// TIA Portal V20 export
// export: Created 2026-10-11T05:19:06.4640986Z, ExportSetting WithDefaults, DisplayName Totally Integrated Automation Portal, DisplayVersion V20, DisplayName TIA Portal Openness, DisplayVersion V20, DisplayName TIA Portal Teamcenter Gateway, DisplayVersion V20, DisplayName TIA Portal Version Control Interface, DisplayVersion V20, DisplayName SINAMICS Startdrive Advanced, DisplayVersion V20 SP1 Update 2, DisplayName SINAMICS Startdrive G110M, G120, G120C, G120D, G120P, G115D, DisplayVersion V20 SP1 Update 2, DisplayName SINAMICS Startdrive G130, G150, S120, S150, SINAMICS MV, G220, S200, S210, DisplayVersion V20 SP1 Update 2, DisplayName STEP 7 Professional, DisplayVersion V20, DisplayName STEP 7 Safety, DisplayVersion V20, DisplayName WinCC Basic/Comfort/Advanced, DisplayVersion V20, DisplayName WinCC Professional, DisplayVersion V20, DisplayName WinCC Unified, DisplayVersion V20
FUNCTION "FRK_Route_InnerUnit" : Bool   // FC65, SCL
{ S7_Optimized_Access := 'TRUE' }
VERSION : 0.1
// stored: AutoNumber true, IsIECCheckEnabled false, SetENOAutomatically false, UDAEnableTagReadback false
   VAR_INPUT
      Request : "ST_HmiRequest";
   END_VAR
   VAR_IN_OUT
      Module : "FB_InnerUnit";
      Hal : "ST_InnerUnitHal";
      Report : "ST_ReleaseReport";
   END_VAR
   VAR_TEMP
      RouteMatched : Bool;
      Index : Int;
   END_VAR
BEGIN

   #FRK_Route_InnerUnit := FALSE;
   IF NOT "FRK_PathOwned"(OwnerPath := #Module.Status.Name, TargetPath := #Request.TargetPath) THEN
       RETURN;
   END_IF;
   "FRK_Release_InnerUnit"(Unit := #Module.Unit,
                           Hal := #Hal);
   "FRK_ManualCommon"(Core := #Module.Core,
                      Unit := #Module.Unit,
                      Status := #Module.Status,
                      Report := #Report);
   IF #Request.TargetPath = STRING_TO_WSTRING(#Module.Status.Name) THEN
       "FRK_ReleaseReason"(Report := #Report,
                           Description := WSTRING#'std.error.unsupportedHmiRequest',
                           Reason := 2008,
                           Path := STRING_TO_WSTRING(#Module.Status.Name),
                           Kind := 4);
       #FRK_Route_InnerUnit := TRUE;
       RETURN;
   END_IF;
   #RouteMatched := "FRK_Route_DeclarationCell"(Module := #Module.Cell, Hal := #Hal.Cell, Request := #Request, Report := #Report);
   #FRK_Route_InnerUnit := #FRK_Route_InnerUnit OR #RouteMatched;
END_FUNCTION
